(* IEC 61131-3 sources: ZPLC/packages/zplc-ide/plant-scenes/merge-lines, 2 files *)

(* ---- reference.st ---- *)
PROGRAM MergeLines
VAR_INPUT
    Start AT %I0.0 : BOOL;
    WaitA AT %I0.1 : BOOL;
    WaitB AT %I0.2 : BOOL;
    Zone  AT %I0.3 : BOOL;
END_VAR
VAR_OUTPUT
    RunA  AT %Q0.0 : BOOL;
    RunB  AT %Q0.1 : BOOL;
    RunOut AT %Q0.2 : BOOL;
    EmitA AT %Q0.3 : BOOL;
    EmitB AT %Q0.4 : BOOL;
    HoldA AT %Q0.5 : BOOL;
    HoldB AT %Q0.6 : BOOL;
    Done  AT %Q0.7 : BOOL;
END_VAR
VAR
    Active : BOOL;
    GrantA : BOOL;
    GrantB : BOOL;
    Seen   : BOOL;
    GoneA  : F_TRIG;
    GoneB  : F_TRIG;
    ZoneGone : F_TRIG;
    LoadedA : CTU;
    LoadedB : CTU;
    Merged  : CTU;
END_VAR

IF Start THEN
    Active := TRUE;
END_IF;

(* each feeder is loaded with three boxes, the next one once the previous has left the blade *)
GoneA(CLK := WaitA);
GoneB(CLK := WaitB);
EmitA := (Start OR GoneA.Q) AND Active AND NOT LoadedA.Q;
EmitB := (Start OR GoneB.Q) AND Active AND NOT LoadedB.Q;
LoadedA(CU := GoneA.Q, R := FALSE, PV := 3);
LoadedB(CU := GoneB.Q, R := FALSE, PV := 3);

(* arbitration: one grant at a time, line A first; a grant ends when its box has left the merge zone *)
ZoneGone(CLK := Zone);
IF Active AND NOT GrantA AND NOT GrantB AND NOT Zone THEN
    IF WaitA THEN
        GrantA := TRUE;
    ELSIF WaitB THEN
        GrantB := TRUE;
    END_IF;
END_IF;
IF (GrantA OR GrantB) AND Zone THEN
    Seen := TRUE;
END_IF;
IF Seen AND ZoneGone.Q THEN
    GrantA := FALSE;
    GrantB := FALSE;
    Seen := FALSE;
END_IF;
Merged(CU := ZoneGone.Q, R := FALSE, PV := 6);

RunA := Active;
RunB := Active;
RunOut := Active;
HoldA := Active AND NOT GrantA;
HoldB := Active AND NOT GrantB;
Done := Merged.Q;

END_PROGRAM

(* ---- starter.st ---- *)
PROGRAM MergeLines
VAR_INPUT
    Start  AT %I0.0 : BOOL;  (* StartButton.pressed: start the line *)
    WaitA  AT %I0.1 : BOOL;  (* EyeA.detect: a box waits at the blade of feeder A *)
    WaitB  AT %I0.2 : BOOL;  (* EyeB.detect: a box waits at the blade of feeder B *)
    Zone   AT %I0.3 : BOOL;  (* EyeZone.detect: a box is on the outfeed past the merge *)
END_VAR
VAR_OUTPUT
    RunA   AT %Q0.0 : BOOL;  (* FeedA.run: run feeder A *)
    RunB   AT %Q0.1 : BOOL;  (* FeedB.run: run feeder B *)
    RunOut AT %Q0.2 : BOOL;  (* Outfeed.run: run the outfeed belt *)
    EmitA  AT %Q0.3 : BOOL;  (* EmitterA.emit: put one box on feeder A *)
    EmitB  AT %Q0.4 : BOOL;  (* EmitterB.emit: put one box on feeder B *)
    HoldA  AT %Q0.5 : BOOL;  (* BladeA.extend: the blade holds feeder A while true *)
    HoldB  AT %Q0.6 : BOOL;  (* BladeB.extend: the blade holds feeder B while true *)
    Done   AT %Q0.7 : BOOL;  (* DoneLight.lit: lit when all six boxes have left *)
END_VAR

(* Goal: a press of the start button loads three boxes on each feeder, one
   at a time, and each blade holds its feeder. Let one box at a time through
   to the outfeed: never open both blades together, and open the next one
   only when the previous box has left the merge, seen at Zone. Light Done
   when all six boxes have left. *)

END_PROGRAM
